Fanuc KAREL source: KT00242.KL

PROGRAM KT00242
%NOLOCKGROUP
VAR
  Y1: ARRAY[2] OF BYTE
  B2: BOOLEAN
  OUT: INTEGER
BEGIN
  Y1[1] = 2
    B2 = FALSE
  OUT = Y1[1] OR B2
END KT00242
